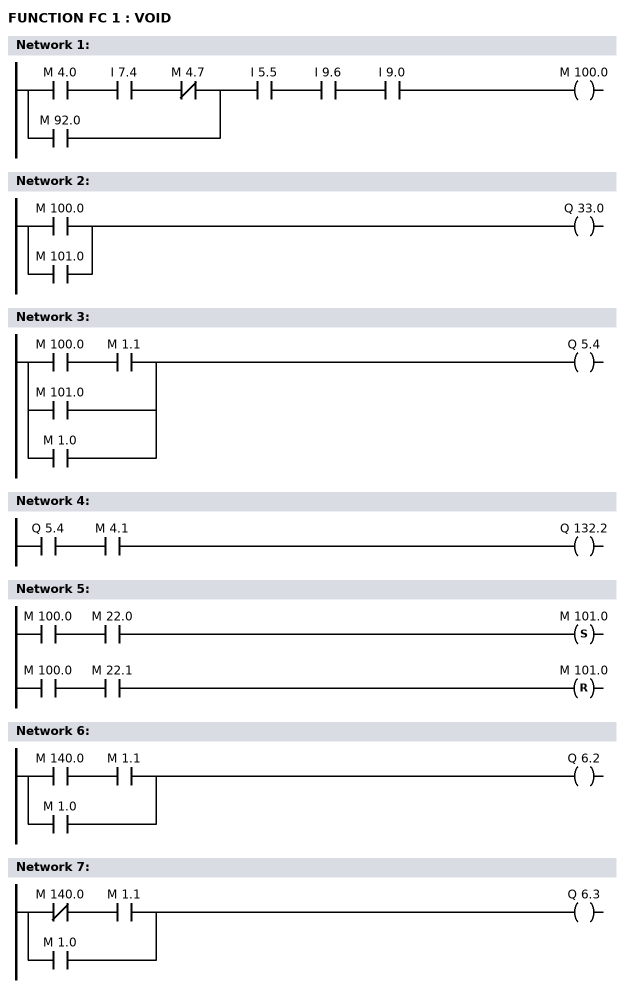

      A(    ;
      A     M      4.0;
      A     I      7.4;
      AN    M      4.7;
      O     M     92.0;
      )     ;
      A     I      5.5;
      A     I      9.6;
      A     I      9.0;
      =     M    100.0;
NETWORK
TITLE =

      O     M    100.0;
      O     M    101.0;
      =     Q     33.0;
NETWORK
TITLE =

      A     M    100.0;
      A     M      1.1;
      O     M    101.0;
      O     M      1.0;
      =     Q      5.4;
NETWORK
TITLE =

      A     Q      5.4;
      A     M      4.1;
      =     Q    132.2;
NETWORK
TITLE =

      A     M    100.0;
      A     M     22.0;
      S     M    101.0;
      A     M    100.0;
      A     M     22.1;
      R     M    101.0;
      NOP   0;
NETWORK
TITLE =

      A     M    140.0;
      A     M      1.1;
      O     M      1.0;
      =     Q      6.2;
NETWORK
TITLE =

      AN    M    140.0;
      A     M      1.1;
      O     M      1.0;
      =     Q      6.3;
NETWORK
TITLE =

      A(    ;
      A     I      8.2;
      L     S5T#150MS;
      SD    T     58;
      NOP   0;
      NOP   0;
      NOP   0;
      A     T     58;
      )     ;
      NOT   ;
      =     Q      7.5;
NETWORK
TITLE =

      A(    ;
      A     I      8.1;
      L     S5T#150MS;
      SD    T     59;
      NOP   0;
      NOP   0;
      NOP   0;
      A     T     59;
      )     ;
      NOT   ;
      =     Q      7.4;
NETWORK
TITLE =
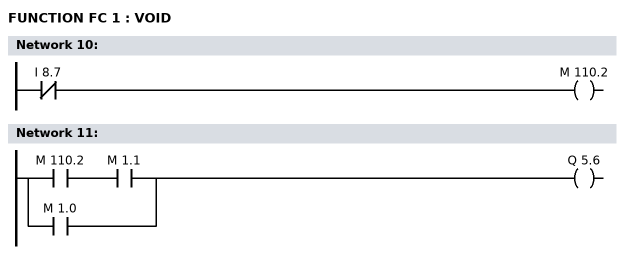

      AN    I      8.7;
      =     M    110.2;
NETWORK
TITLE =

      A     M    110.2;
      A     M      1.1;
      O     M      1.0;
      =     Q      5.6;
NETWORK
TITLE =

      O(    ;
      A     I      8.0;
      L     S5T#150MS;
      SD    T     50;
      NOP   0;
      NOP   0;
      NOP   0;
      A     T     50;
      )     ;
      O     M      1.0;
      =     Q      5.0;
NETWORK
TITLE =
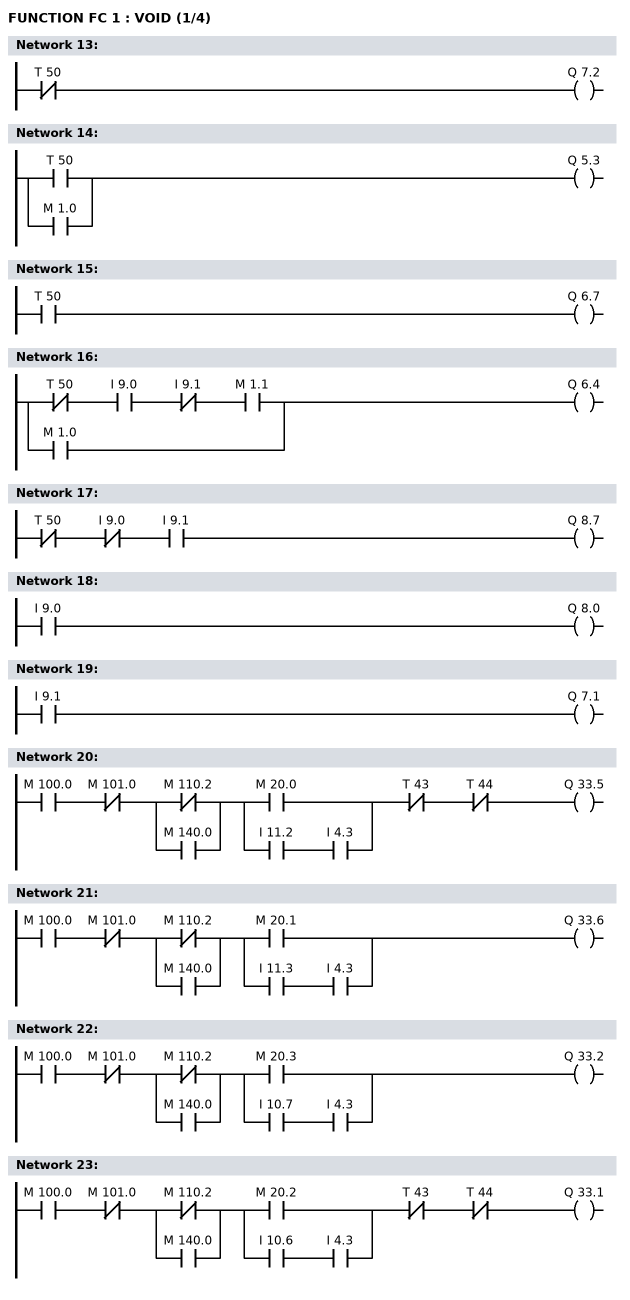

      AN    T     50;
      =     Q      7.2;
NETWORK
TITLE =

      O     T     50;
      O     M      1.0;
      =     Q      5.3;
NETWORK
TITLE =

      A     T     50;
      =     Q      6.7;
NETWORK
TITLE =

      AN    T     50;
      A     I      9.0;
      AN    I      9.1;
      A     M      1.1;
      O     M      1.0;
      =     Q      6.4;
NETWORK
TITLE =

      AN    T     50;
      AN    I      9.0;
      A     I      9.1;
      =     Q      8.7;
NETWORK
TITLE =

      A     I      9.0;
      =     Q      8.0;
NETWORK
TITLE =

      A     I      9.1;
      =     Q      7.1;
NETWORK
TITLE =

      A     M    100.0;
      AN    M    101.0;
      A(    ;
      ON    M    110.2;
      O     M    140.0;
      )     ;
      A(    ;
      O     M     20.0;
      O     ;
      A     I     11.2;
      A     I      4.3;
      )     ;
      AN    T     43;
      AN    T     44;
      =     Q     33.5;
NETWORK
TITLE =

      A     M    100.0;
      AN    M    101.0;
      A(    ;
      ON    M    110.2;
      O     M    140.0;
      )     ;
      A(    ;
      O     M     20.1;
      O     ;
      A     I     11.3;
      A     I      4.3;
      )     ;
      =     Q     33.6;
NETWORK
TITLE =

      A     M    100.0;
      AN    M    101.0;
      A(    ;
      ON    M    110.2;
      O     M    140.0;
      )     ;
      A(    ;
      O     M     20.3;
      O     ;
      A     I     10.7;
      A     I      4.3;
      )     ;
      =     Q     33.2;
NETWORK
TITLE =

      A     M    100.0;
      AN    M    101.0;
      A(    ;
      ON    M    110.2;
      O     M    140.0;
      )     ;
      A(    ;
      O     M     20.2;
      O     ;
      A     I     10.6;
      A     I      4.3;
      )     ;
      AN    T     43;
      AN    T     44;
      =     Q     33.1;
NETWORK
TITLE =
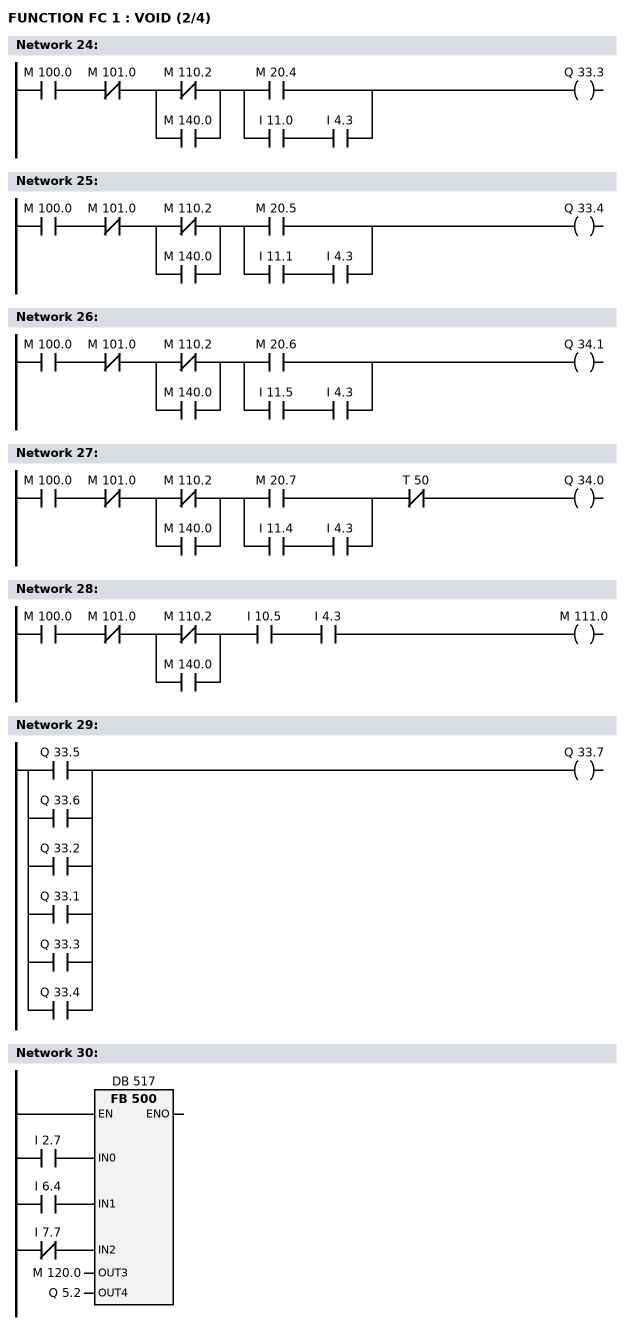

      A     M    100.0;
      AN    M    101.0;
      A(    ;
      ON    M    110.2;
      O     M    140.0;
      )     ;
      A(    ;
      O     M     20.4;
      O     ;
      A     I     11.0;
      A     I      4.3;
      )     ;
      =     Q     33.3;
NETWORK
TITLE =

      A     M    100.0;
      AN    M    101.0;
      A(    ;
      ON    M    110.2;
      O     M    140.0;
      )     ;
      A(    ;
      O     M     20.5;
      O     ;
      A     I     11.1;
      A     I      4.3;
      )     ;
      =     Q     33.4;
NETWORK
TITLE =

      A     M    100.0;
      AN    M    101.0;
      A(    ;
      ON    M    110.2;
      O     M    140.0;
      )     ;
      A(    ;
      O     M     20.6;
      O     ;
      A     I     11.5;
      A     I      4.3;
      )     ;
      =     Q     34.1;
NETWORK
TITLE =

      A     M    100.0;
      AN    M    101.0;
      A(    ;
      ON    M    110.2;
      O     M    140.0;
      )     ;
      A(    ;
      O     M     20.7;
      O     ;
      A     I     11.4;
      A     I      4.3;
      )     ;
      AN    T     50;
      =     Q     34.0;
NETWORK
TITLE =

      A     M    100.0;
      AN    M    101.0;
      A(    ;
      ON    M    110.2;
      O     M    140.0;
      )     ;
      A     I     10.5;
      A     I      4.3;
      =     M    111.0;
NETWORK
TITLE =

      O     Q     33.5;
      O     Q     33.6;
      O     Q     33.2;
      O     Q     33.1;
      O     Q     33.3;
      O     Q     33.4;
      =     Q     33.7;
NETWORK
TITLE =

      A     I      2.7;
      =     L      0.0;
      BLD   103;
      A     I      6.4;
      =     L      0.1;
      BLD   103;
      AN    I      7.7;
      =     L      0.2;
      BLD   103;
      CALL FB   500 , DB   517 (
           IN0                      := L      0.0,
           IN1                      := L      0.1,
           IN2                      := L      0.2,
           OUT3                     := M    120.0,
           OUT4                     := Q      5.2);
      NOP   0;
NETWORK
TITLE =
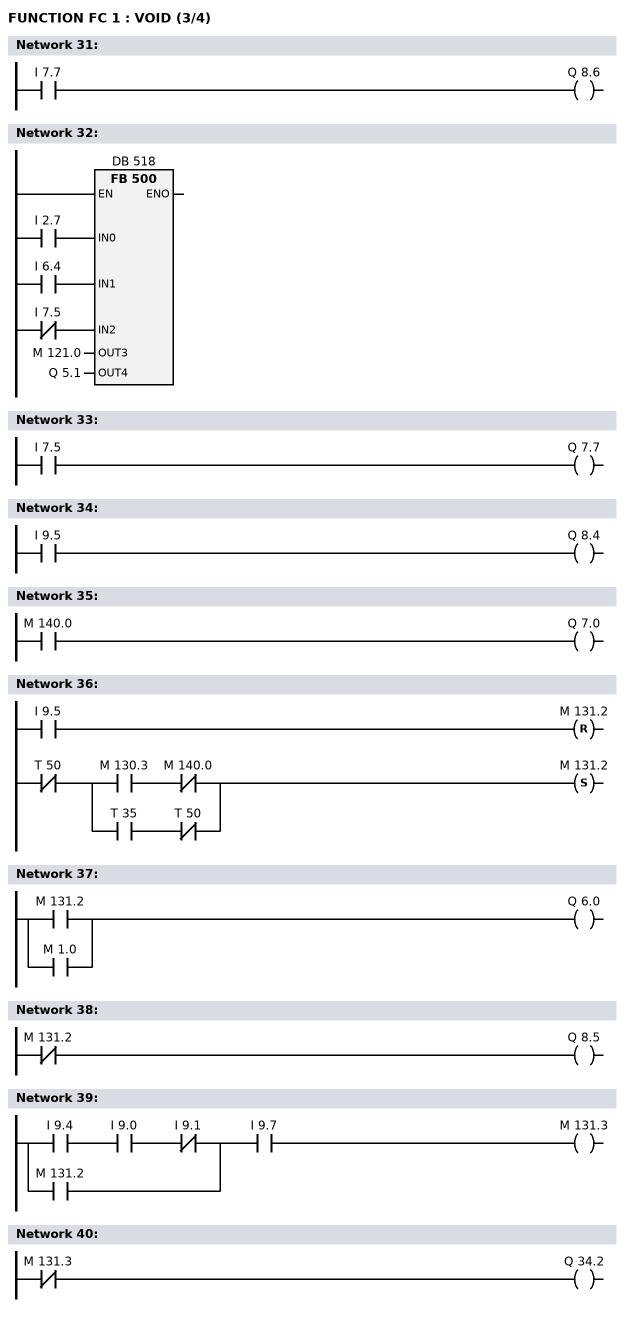

      A     I      7.7;
      =     Q      8.6;
NETWORK
TITLE =

      A     I      2.7;
      =     L      0.0;
      BLD   103;
      A     I      6.4;
      =     L      0.1;
      BLD   103;
      AN    I      7.5;
      =     L      0.2;
      BLD   103;
      CALL FB   500 , DB   518 (
           IN0                      := L      0.0,
           IN1                      := L      0.1,
           IN2                      := L      0.2,
           OUT3                     := M    121.0,
           OUT4                     := Q      5.1);
      NOP   0;
NETWORK
TITLE =

      A     I      7.5;
      =     Q      7.7;
NETWORK
TITLE =

      A     I      9.5;
      =     Q      8.4;
NETWORK
TITLE =

      A     M    140.0;
      =     Q      7.0;
NETWORK
TITLE =

      A     I      9.5;
      R     M    131.2;
      AN    T     50;
      A(    ;
      A     M    130.3;
      AN    M    140.0;
      O     ;
      A     T     35;
      AN    T     50;
      )     ;
      S     M    131.2;
      NOP   0;
NETWORK
TITLE =

      O     M    131.2;
      O     M      1.0;
      =     Q      6.0;
NETWORK
TITLE =

      AN    M    131.2;
      =     Q      8.5;
NETWORK
TITLE =

      A(    ;
      A     I      9.4;
      A     I      9.0;
      AN    I      9.1;
      O     M    131.2;
      )     ;
      A     I      9.7;
      =     M    131.3;
NETWORK
TITLE =

      AN    M    131.3;
      =     Q     34.2;
NETWORK
TITLE =
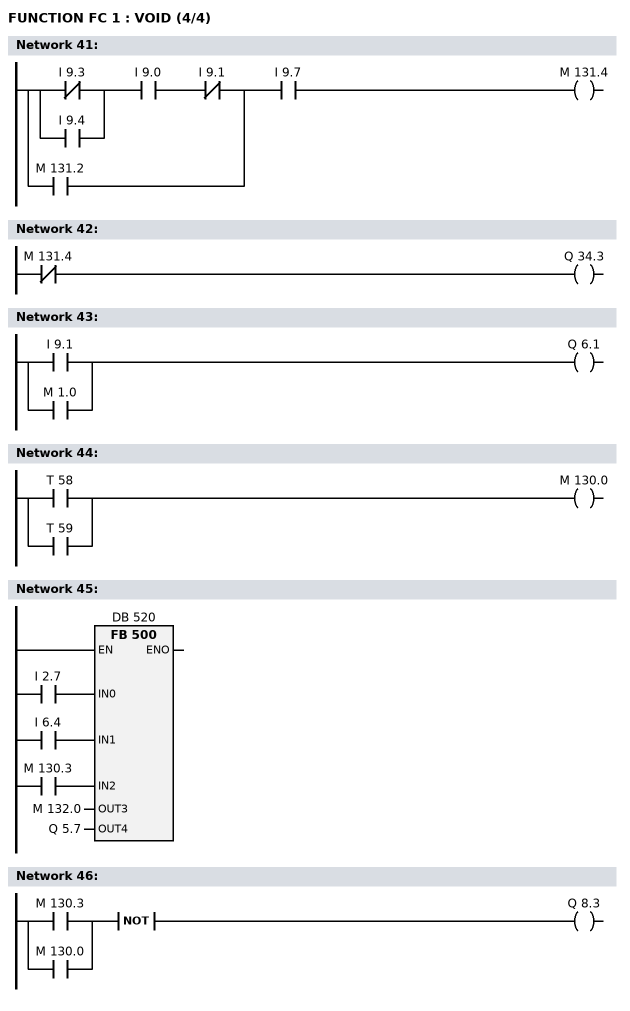

      A(    ;
      A(    ;
      ON    I      9.3;
      O     I      9.4;
      )     ;
      A     I      9.0;
      AN    I      9.1;
      O     M    131.2;
      )     ;
      A     I      9.7;
      =     M    131.4;
NETWORK
TITLE =

      AN    M    131.4;
      =     Q     34.3;
NETWORK
TITLE =

      O     I      9.1;
      O     M      1.0;
      =     Q      6.1;
NETWORK
TITLE =

      O     T     58;
      O     T     59;
      =     M    130.0;
NETWORK
TITLE =

      A     I      2.7;
      =     L      0.0;
      BLD   103;
      A     I      6.4;
      =     L      0.1;
      BLD   103;
      A     M    130.3;
      =     L      0.2;
      BLD   103;
      CALL FB   500 , DB   520 (
           IN0                      := L      0.0,
           IN1                      := L      0.1,
           IN2                      := L      0.2,
           OUT3                     := M    132.0,
           OUT4                     := Q      5.7);
      NOP   0;
NETWORK
TITLE =

      A(    ;
      O     M    130.3;
      O     M    130.0;
      )     ;
      NOT   ;
      =     Q      8.3;
NETWORK
TITLE =

      A(    ;
      A     I      8.4;
      L     S5T#150MS;
      SD    T     43;
      NOP   0;
      NOP   0;
      NOP   0;
      A     T     43;
      )     ;
      NOT   ;
      =     Q      6.6;
NETWORK
TITLE =

      A(    ;
      A     I      8.6;
      L     S5T#150MS;
      SD    T     44;
      NOP   0;
      NOP   0;
      NOP   0;
      A     T     44;
      )     ;
      NOT   ;
      =     Q      8.1;
NETWORK
TITLE =

      A(    ;
      A     I      8.5;
      L     S5T#150MS;
      SD    T     46;
      NOP   0;
      NOP   0;
      NOP   0;
      A     T     46;
      )     ;
      NOT   ;
      =     Q      7.6;
NETWORK
TITLE =

      A(    ;
      A     I      8.3;
      L     S5T#150MS;
      SD    T     47;
      NOP   0;
      NOP   0;
      NOP   0;
      A     T     47;
      )     ;
      NOT   ;
      =     Q      8.2;
NETWORK
TITLE =
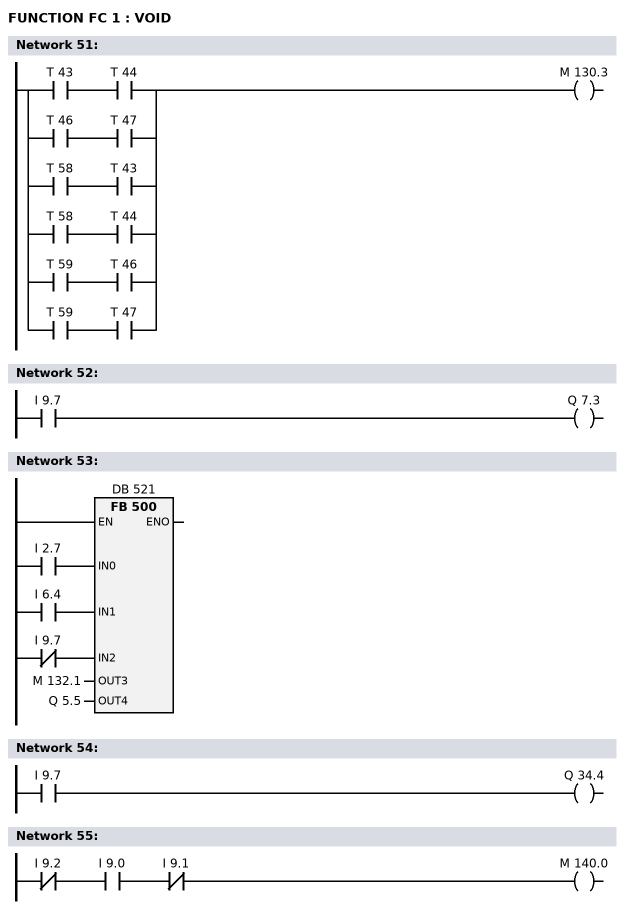

      A     T     43;
      A     T     44;
      O     ;
      A     T     46;
      A     T     47;
      O     ;
      A     T     58;
      A     T     43;
      O     ;
      A     T     58;
      A     T     44;
      O     ;
      A     T     59;
      A     T     46;
      O     ;
      A     T     59;
      A     T     47;
      =     M    130.3;
NETWORK
TITLE =

      A     I      9.7;
      =     Q      7.3;
NETWORK
TITLE =

      A     I      2.7;
      =     L      0.0;
      BLD   103;
      A     I      6.4;
      =     L      0.1;
      BLD   103;
      AN    I      9.7;
      =     L      0.2;
      BLD   103;
      CALL FB   500 , DB   521 (
           IN0                      := L      0.0,
           IN1                      := L      0.1,
           IN2                      := L      0.2,
           OUT3                     := M    132.1,
           OUT4                     := Q      5.5);
      NOP   0;
NETWORK
TITLE =

      A     I      9.7;
      =     Q     34.4;
NETWORK
TITLE =

      AN    I      9.2;
      A     I      9.0;
      AN    I      9.1;
      =     M    140.0;
END_FUNCTION

FUNCTION FC 2 : VOID
VERSION : 0.1

BEGIN
NETWORK
TITLE =
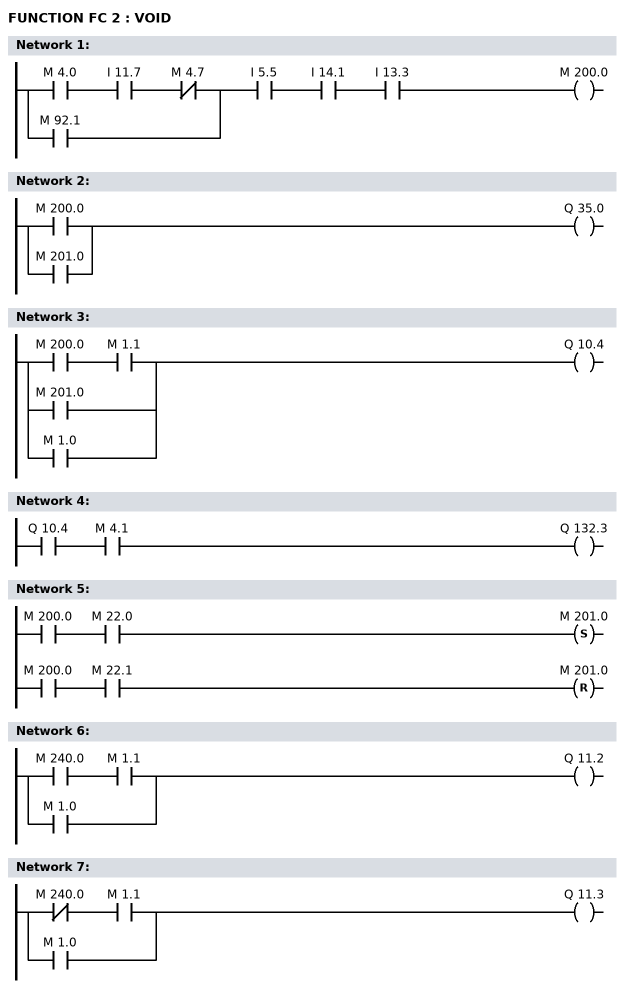

      A(    ;
      A     M      4.0;
      A     I     11.7;
      AN    M      4.7;
      O     M     92.1;
      )     ;
      A     I      5.5;
      A     I     14.1;
      A     I     13.3;
      =     M    200.0;
NETWORK
TITLE =

      O     M    200.0;
      O     M    201.0;
      =     Q     35.0;
NETWORK
TITLE =

      A     M    200.0;
      A     M      1.1;
      O     M    201.0;
      O     M      1.0;
      =     Q     10.4;
NETWORK
TITLE =

      A     Q     10.4;
      A     M      4.1;
      =     Q    132.3;
NETWORK
TITLE =

      A     M    200.0;
      A     M     22.0;
      S     M    201.0;
      A     M    200.0;
      A     M     22.1;
      R     M    201.0;
      NOP   0;
NETWORK
TITLE =

      A     M    240.0;
      A     M      1.1;
      O     M      1.0;
      =     Q     11.2;
NETWORK
TITLE =

      AN    M    240.0;
      A     M      1.1;
      O     M      1.0;
      =     Q     11.3;
NETWORK
TITLE =

      A(    ;
      A     I     12.5;
      L     S5T#150MS;
      SD    T     78;
      NOP   0;
      NOP   0;
      NOP   0;
      A     T     78;
      )     ;
      NOT   ;
      =     Q     12.5;
NETWORK
TITLE =

      A(    ;
      A     I     12.4;
      L     S5T#150MS;
      SD    T     79;
      NOP   0;
      NOP   0;
      NOP   0;
      A     T     79;
      )     ;
      NOT   ;
      =     Q     12.4;
NETWORK
TITLE =
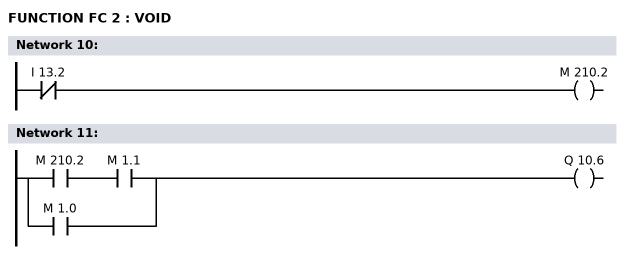

      AN    I     13.2;
      =     M    210.2;
NETWORK
TITLE =

      A     M    210.2;
      A     M      1.1;
      O     M      1.0;
      =     Q     10.6;
NETWORK
TITLE =

      O(    ;
      A     I     12.3;
      L     S5T#150MS;
      SD    T     70;
      NOP   0;
      NOP   0;
      NOP   0;
      A     T     70;
      )     ;
      O     M      1.0;
      =     Q     10.0;
NETWORK
TITLE =
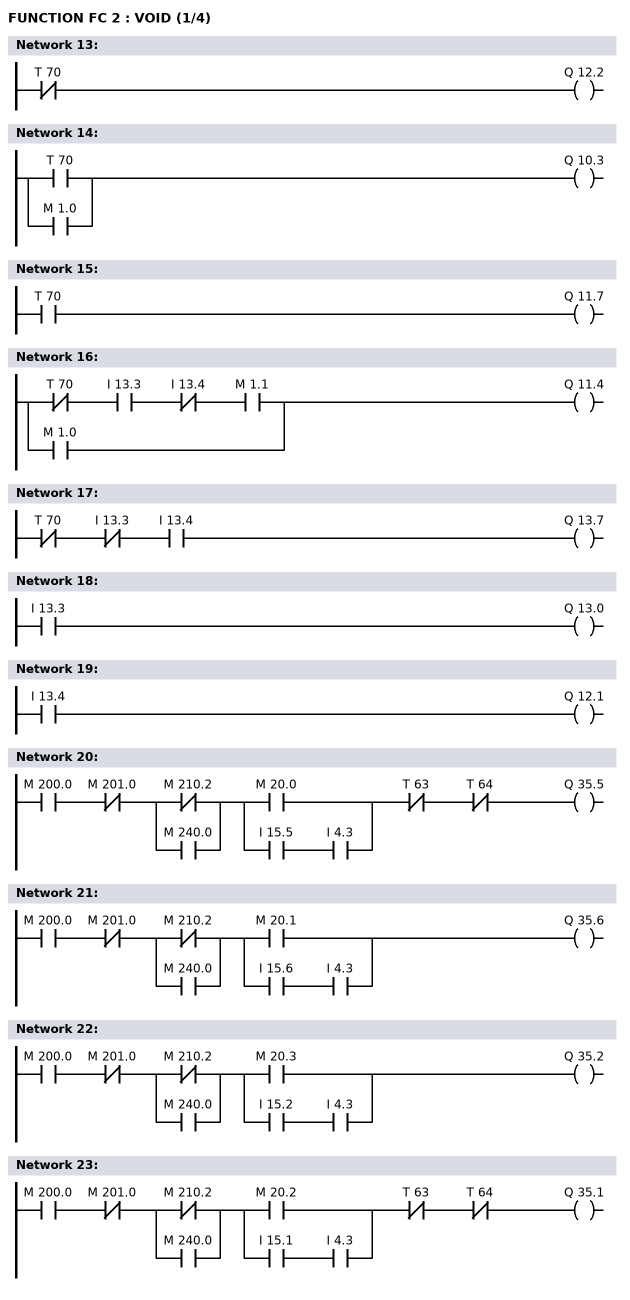

      AN    T     70;
      =     Q     12.2;
NETWORK
TITLE =

      O     T     70;
      O     M      1.0;
      =     Q     10.3;
NETWORK
TITLE =

      A     T     70;
      =     Q     11.7;
NETWORK
TITLE =

      AN    T     70;
      A     I     13.3;
      AN    I     13.4;
      A     M      1.1;
      O     M      1.0;
      =     Q     11.4;
NETWORK
TITLE =

      AN    T     70;
      AN    I     13.3;
      A     I     13.4;
      =     Q     13.7;
NETWORK
TITLE =

      A     I     13.3;
      =     Q     13.0;
NETWORK
TITLE =

      A     I     13.4;
      =     Q     12.1;
NETWORK
TITLE =

      A     M    200.0;
      AN    M    201.0;
      A(    ;
      ON    M    210.2;
      O     M    240.0;
      )     ;
      A(    ;
      O     M     20.0;
      O     ;
      A     I     15.5;
      A     I      4.3;
      )     ;
      AN    T     63;
      AN    T     64;
      =     Q     35.5;
NETWORK
TITLE =

      A     M    200.0;
      AN    M    201.0;
      A(    ;
      ON    M    210.2;
      O     M    240.0;
      )     ;
      A(    ;
      O     M     20.1;
      O     ;
      A     I     15.6;
      A     I      4.3;
      )     ;
      =     Q     35.6;
NETWORK
TITLE =

      A     M    200.0;
      AN    M    201.0;
      A(    ;
      ON    M    210.2;
      O     M    240.0;
      )     ;
      A(    ;
      O     M     20.3;
      O     ;
      A     I     15.2;
      A     I      4.3;
      )     ;
      =     Q     35.2;
NETWORK
TITLE =

      A     M    200.0;
      AN    M    201.0;
      A(    ;
      ON    M    210.2;
      O     M    240.0;
      )     ;
      A(    ;
      O     M     20.2;
      O     ;
      A     I     15.1;
      A     I      4.3;
      )     ;
      AN    T     63;
      AN    T     64;
      =     Q     35.1;
NETWORK
TITLE =
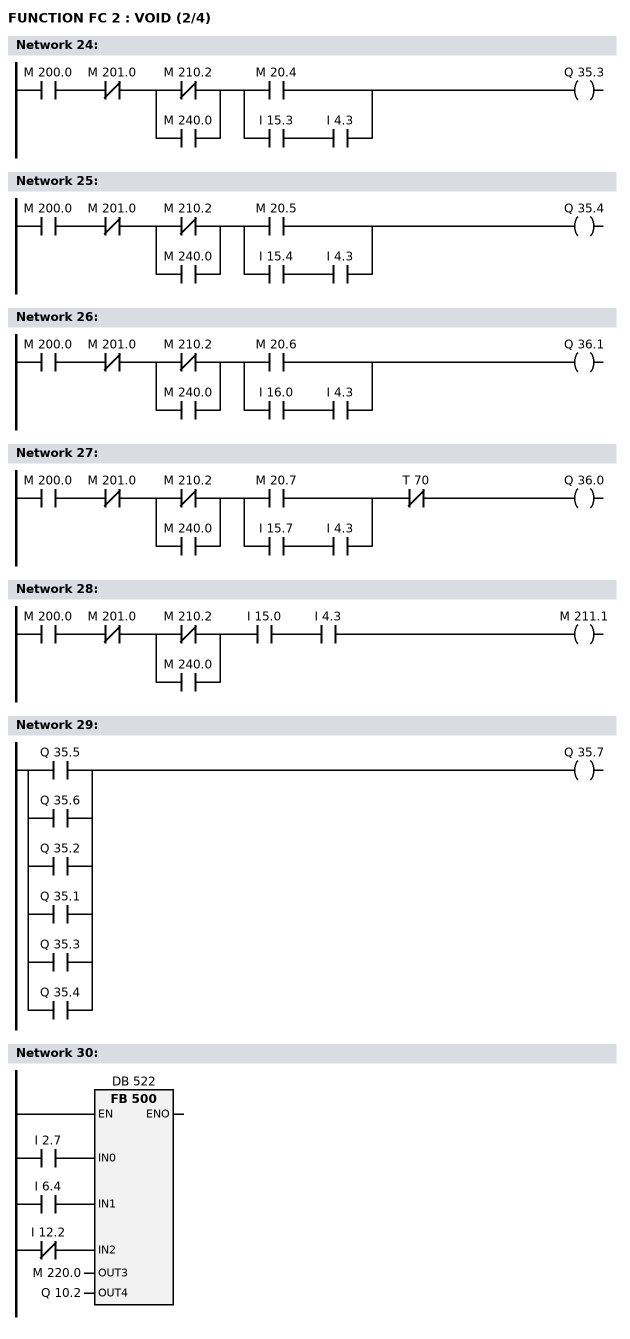

      A     M    200.0;
      AN    M    201.0;
      A(    ;
      ON    M    210.2;
      O     M    240.0;
      )     ;
      A(    ;
      O     M     20.4;
      O     ;
      A     I     15.3;
      A     I      4.3;
      )     ;
      =     Q     35.3;
NETWORK
TITLE =

      A     M    200.0;
      AN    M    201.0;
      A(    ;
      ON    M    210.2;
      O     M    240.0;
      )     ;
      A(    ;
      O     M     20.5;
      O     ;
      A     I     15.4;
      A     I      4.3;
      )     ;
      =     Q     35.4;
NETWORK
TITLE =

      A     M    200.0;
      AN    M    201.0;
      A(    ;
      ON    M    210.2;
      O     M    240.0;
      )     ;
      A(    ;
      O     M     20.6;
      O     ;
      A     I     16.0;
      A     I      4.3;
      )     ;
      =     Q     36.1;
NETWORK
TITLE =

      A     M    200.0;
      AN    M    201.0;
      A(    ;
      ON    M    210.2;
      O     M    240.0;
      )     ;
      A(    ;
      O     M     20.7;
      O     ;
      A     I     15.7;
      A     I      4.3;
      )     ;
      AN    T     70;
      =     Q     36.0;
NETWORK
TITLE =

      A     M    200.0;
      AN    M    201.0;
      A(    ;
      ON    M    210.2;
      O     M    240.0;
      )     ;
      A     I     15.0;
      A     I      4.3;
      =     M    211.1;
NETWORK
TITLE =

      O     Q     35.5;
      O     Q     35.6;
      O     Q     35.2;
      O     Q     35.1;
      O     Q     35.3;
      O     Q     35.4;
      =     Q     35.7;
NETWORK
TITLE =

      A     I      2.7;
      =     L      0.0;
      BLD   103;
      A     I      6.4;
      =     L      0.1;
      BLD   103;
      AN    I     12.2;
      =     L      0.2;
      BLD   103;
      CALL FB   500 , DB   522 (
           IN0                      := L      0.0,
           IN1                      := L      0.1,
           IN2                      := L      0.2,
           OUT3                     := M    220.0,
           OUT4                     := Q     10.2);
      NOP   0;
NETWORK
TITLE =
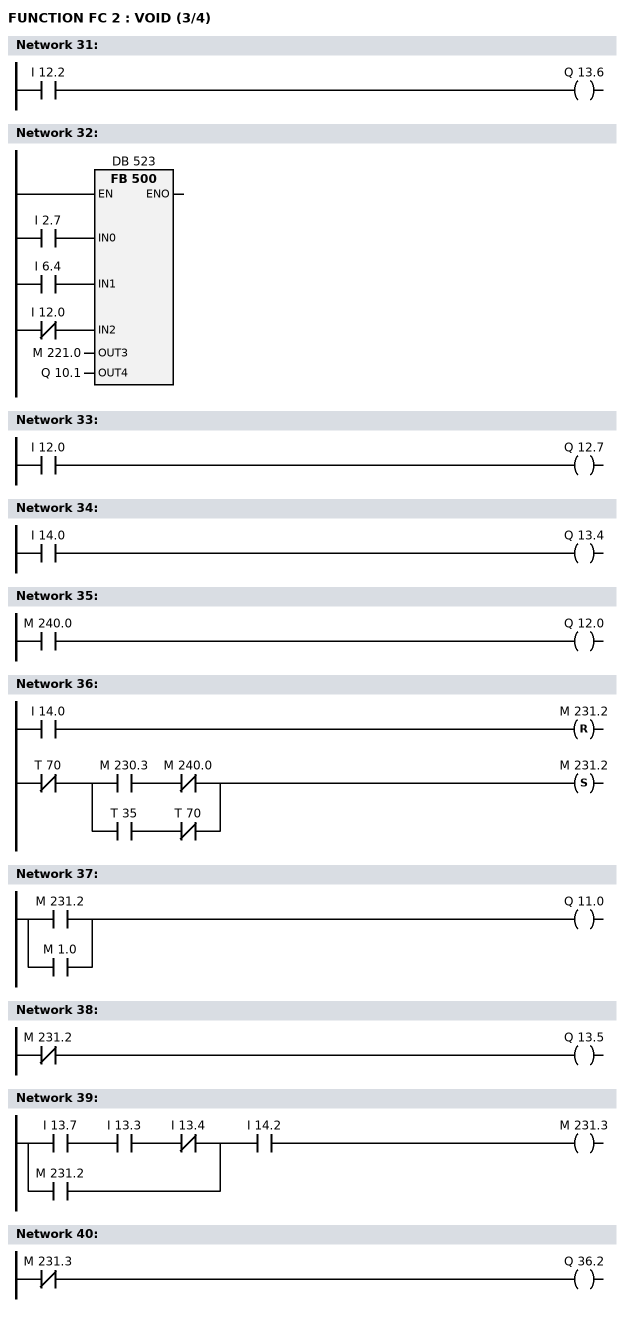

      A     I     12.2;
      =     Q     13.6;
NETWORK
TITLE =

      A     I      2.7;
      =     L      0.0;
      BLD   103;
      A     I      6.4;
      =     L      0.1;
      BLD   103;
      AN    I     12.0;
      =     L      0.2;
      BLD   103;
      CALL FB   500 , DB   523 (
           IN0                      := L      0.0,
           IN1                      := L      0.1,
           IN2                      := L      0.2,
           OUT3                     := M    221.0,
           OUT4                     := Q     10.1);
      NOP   0;
NETWORK
TITLE =

      A     I     12.0;
      =     Q     12.7;
NETWORK
TITLE =

      A     I     14.0;
      =     Q     13.4;
NETWORK
TITLE =

      A     M    240.0;
      =     Q     12.0;
NETWORK
TITLE =

      A     I     14.0;
      R     M    231.2;
      AN    T     70;
      A(    ;
      A     M    230.3;
      AN    M    240.0;
      O     ;
      A     T     35;
      AN    T     70;
      )     ;
      S     M    231.2;
      NOP   0;
NETWORK
TITLE =

      O     M    231.2;
      O     M      1.0;
      =     Q     11.0;
NETWORK
TITLE =

      AN    M    231.2;
      =     Q     13.5;
NETWORK
TITLE =

      A(    ;
      A     I     13.7;
      A     I     13.3;
      AN    I     13.4;
      O     M    231.2;
      )     ;
      A     I     14.2;
      =     M    231.3;
NETWORK
TITLE =

      AN    M    231.3;
      =     Q     36.2;
NETWORK
TITLE =
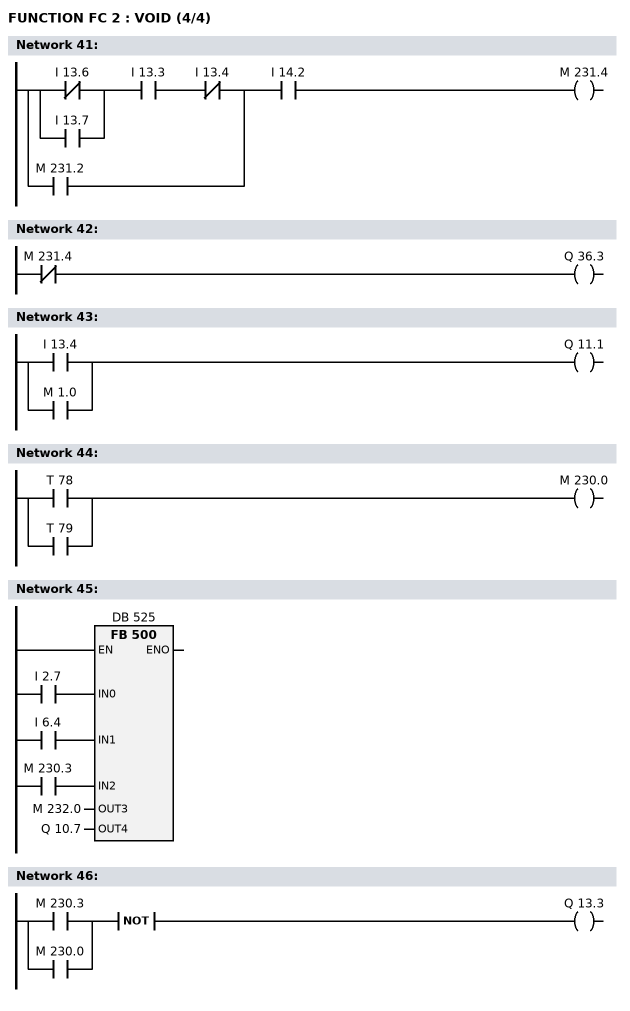

      A(    ;
      A(    ;
      ON    I     13.6;
      O     I     13.7;
      )     ;
      A     I     13.3;
      AN    I     13.4;
      O     M    231.2;
      )     ;
      A     I     14.2;
      =     M    231.4;
NETWORK
TITLE =

      AN    M    231.4;
      =     Q     36.3;
NETWORK
TITLE =

      O     I     13.4;
      O     M      1.0;
      =     Q     11.1;
NETWORK
TITLE =

      O     T     78;
      O     T     79;
      =     M    230.0;
NETWORK
TITLE =

      A     I      2.7;
      =     L      0.0;
      BLD   103;
      A     I      6.4;
      =     L      0.1;
      BLD   103;
      A     M    230.3;
      =     L      0.2;
      BLD   103;
      CALL FB   500 , DB   525 (
           IN0                      := L      0.0,
           IN1                      := L      0.1,
           IN2                      := L      0.2,
           OUT3                     := M    232.0,
           OUT4                     := Q     10.7);
      NOP   0;
NETWORK
TITLE =

      A(    ;
      O     M    230.3;
      O     M    230.0;
      )     ;
      NOT   ;
      =     Q     13.3;
NETWORK
TITLE =

      A(    ;
      A     I     12.7;
      L     S5T#150MS;
      SD    T     63;
      NOP   0;
      NOP   0;
      NOP   0;
      A     T     63;
      )     ;
      NOT   ;
      =     Q     11.6;
NETWORK
TITLE =

      A(    ;
      A     I     13.1;
      L     S5T#150MS;
      SD    T     64;
      NOP   0;
      NOP   0;
      NOP   0;
      A     T     64;
      )     ;
      NOT   ;
      =     Q     13.1;
NETWORK
TITLE =

      A(    ;
      A     I     13.0;
      L     S5T#150MS;
      SD    T     66;
      NOP   0;
      NOP   0;
      NOP   0;
      A     T     66;
      )     ;
      NOT   ;
      =     Q     12.6;
NETWORK
TITLE =

      A(    ;
      A     I     12.6;
      L     S5T#150MS;
      SD    T     67;
      NOP   0;
      NOP   0;
      NOP   0;
      A     T     67;
      )     ;
      NOT   ;
      =     Q     13.2;
NETWORK
TITLE =
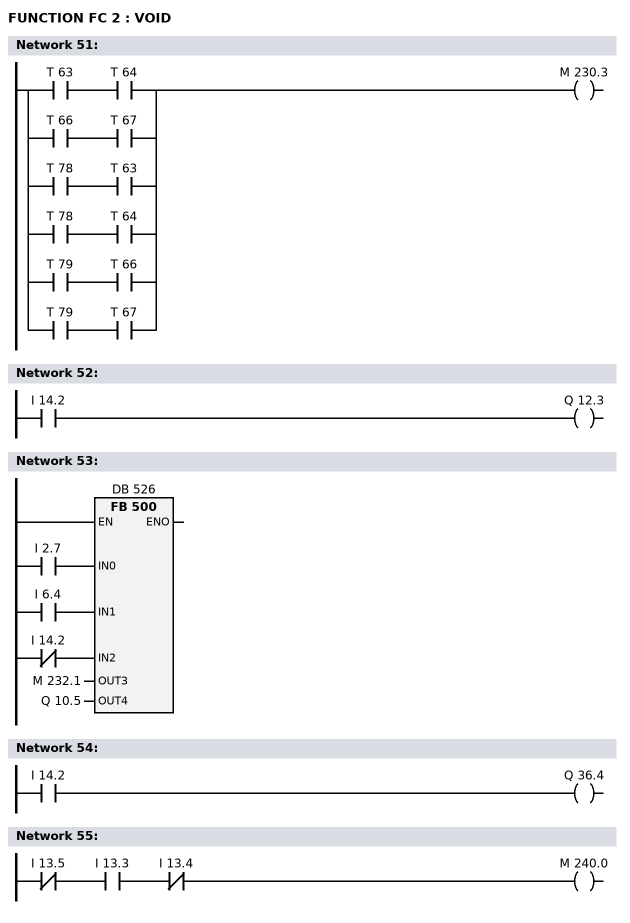

      A     T     63;
      A     T     64;
      O     ;
      A     T     66;
      A     T     67;
      O     ;
      A     T     78;
      A     T     63;
      O     ;
      A     T     78;
      A     T     64;
      O     ;
      A     T     79;
      A     T     66;
      O     ;
      A     T     79;
      A     T     67;
      =     M    230.3;
NETWORK
TITLE =

      A     I     14.2;
      =     Q     12.3;
NETWORK
TITLE =

      A     I      2.7;
      =     L      0.0;
      BLD   103;
      A     I      6.4;
      =     L      0.1;
      BLD   103;
      AN    I     14.2;
      =     L      0.2;
      BLD   103;
      CALL FB   500 , DB   526 (
           IN0                      := L      0.0,
           IN1                      := L      0.1,
           IN2                      := L      0.2,
           OUT3                     := M    232.1,
           OUT4                     := Q     10.5);
      NOP   0;
NETWORK
TITLE =

      A     I     14.2;
      =     Q     36.4;
NETWORK
TITLE =

      AN    I     13.5;
      A     I     13.3;
      AN    I     13.4;
      =     M    240.0;
END_FUNCTION

FUNCTION FC 3 : VOID
VERSION : 0.1

BEGIN
NETWORK
TITLE =
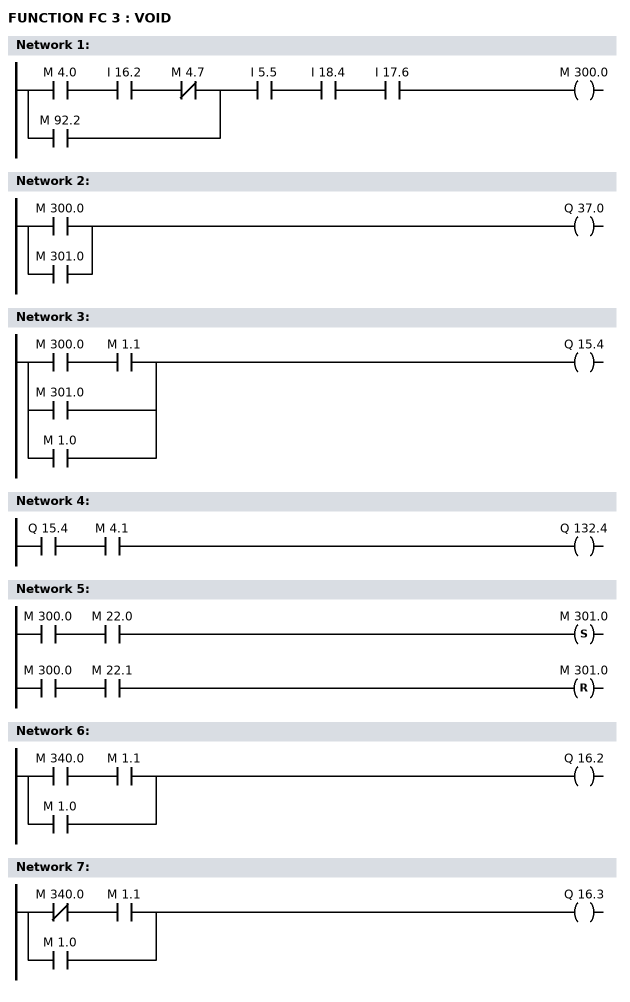

      A(    ;
      A     M      4.0;
      A     I     16.2;
      AN    M      4.7;
      O     M     92.2;
      )     ;
      A     I      5.5;
      A     I     18.4;
      A     I     17.6;
      =     M    300.0;
NETWORK
TITLE =

      O     M    300.0;
      O     M    301.0;
      =     Q     37.0;
NETWORK
TITLE =

      A     M    300.0;
      A     M      1.1;
      O     M    301.0;
      O     M      1.0;
      =     Q     15.4;
NETWORK
TITLE =

      A     Q     15.4;
      A     M      4.1;
      =     Q    132.4;
NETWORK
TITLE =

      A     M    300.0;
      A     M     22.0;
      S     M    301.0;
      A     M    300.0;
      A     M     22.1;
      R     M    301.0;
      NOP   0;
NETWORK
TITLE =

      A     M    340.0;
      A     M      1.1;
      O     M      1.0;
      =     Q     16.2;
NETWORK
TITLE =

      AN    M    340.0;
      A     M      1.1;
      O     M      1.0;
      =     Q     16.3;
NETWORK
TITLE =

      A(    ;
      A     I     17.0;
      L     S5T#150MS;
      SD    T     98;
      NOP   0;
      NOP   0;
      NOP   0;
      A     T     98;
      )     ;
      NOT   ;
      =     Q     17.5;
NETWORK
TITLE =

      A(    ;
      A     I     16.7;
      L     S5T#150MS;
      SD    T     99;
      NOP   0;
      NOP   0;
      NOP   0;
      A     T     99;
      )     ;
      NOT   ;
      =     Q     17.4;
NETWORK
TITLE =
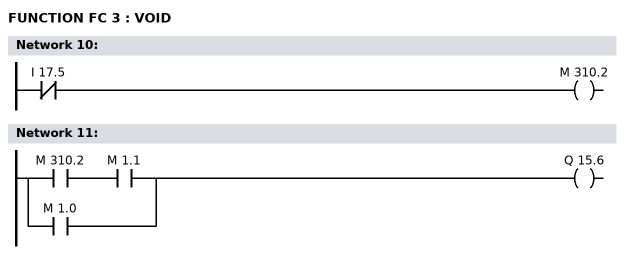

      AN    I     17.5;
      =     M    310.2;
NETWORK
TITLE =

      A     M    310.2;
      A     M      1.1;
      O     M      1.0;
      =     Q     15.6;
NETWORK
TITLE =

      O(    ;
      A     I     16.6;
      L     S5T#150MS;
      SD    T     90;
      NOP   0;
      NOP   0;
      NOP   0;
      A     T     90;
      )     ;
      O     M      1.0;
      =     Q     15.0;
NETWORK
TITLE =
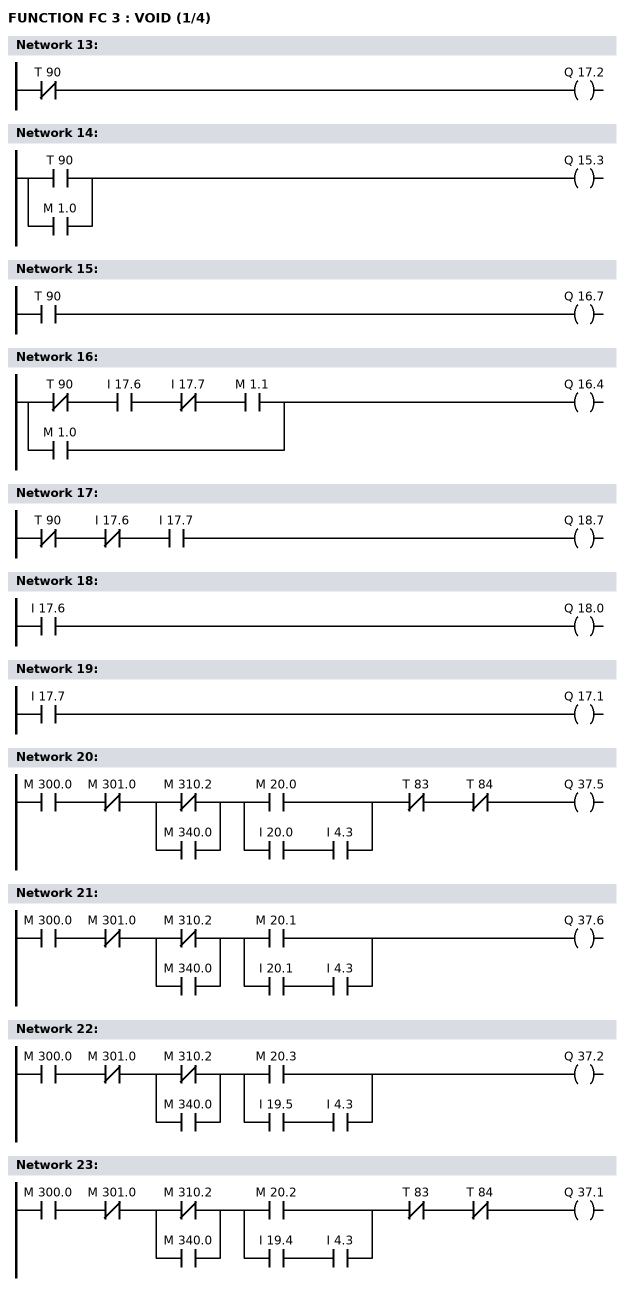

      AN    T     90;
      =     Q     17.2;
NETWORK
TITLE =

      O     T     90;
      O     M      1.0;
      =     Q     15.3;
NETWORK
TITLE =

      A     T     90;
      =     Q     16.7;
NETWORK
TITLE =

      AN    T     90;
      A     I     17.6;
      AN    I     17.7;
      A     M      1.1;
      O     M      1.0;
      =     Q     16.4;
NETWORK
TITLE =

      AN    T     90;
      AN    I     17.6;
      A     I     17.7;
      =     Q     18.7;
NETWORK
TITLE =

      A     I     17.6;
      =     Q     18.0;
NETWORK
TITLE =

      A     I     17.7;
      =     Q     17.1;
NETWORK
TITLE =

      A     M    300.0;
      AN    M    301.0;
      A(    ;
      ON    M    310.2;
      O     M    340.0;
      )     ;
      A(    ;
      O     M     20.0;
      O     ;
      A     I     20.0;
      A     I      4.3;
      )     ;
      AN    T     83;
      AN    T     84;
      =     Q     37.5;
NETWORK
TITLE =

      A     M    300.0;
      AN    M    301.0;
      A(    ;
      ON    M    310.2;
      O     M    340.0;
      )     ;
      A(    ;
      O     M     20.1;
      O     ;
      A     I     20.1;
      A     I      4.3;
      )     ;
      =     Q     37.6;
NETWORK
TITLE =

      A     M    300.0;
      AN    M    301.0;
      A(    ;
      ON    M    310.2;
      O     M    340.0;
      )     ;
      A(    ;
      O     M     20.3;
      O     ;
      A     I     19.5;
      A     I      4.3;
      )     ;
      =     Q     37.2;
NETWORK
TITLE =

      A     M    300.0;
      AN    M    301.0;
      A(    ;
      ON    M    310.2;
      O     M    340.0;
      )     ;
      A(    ;
      O     M     20.2;
      O     ;
      A     I     19.4;
      A     I      4.3;
      )     ;
      AN    T     83;
      AN    T     84;
      =     Q     37.1;
NETWORK
TITLE =
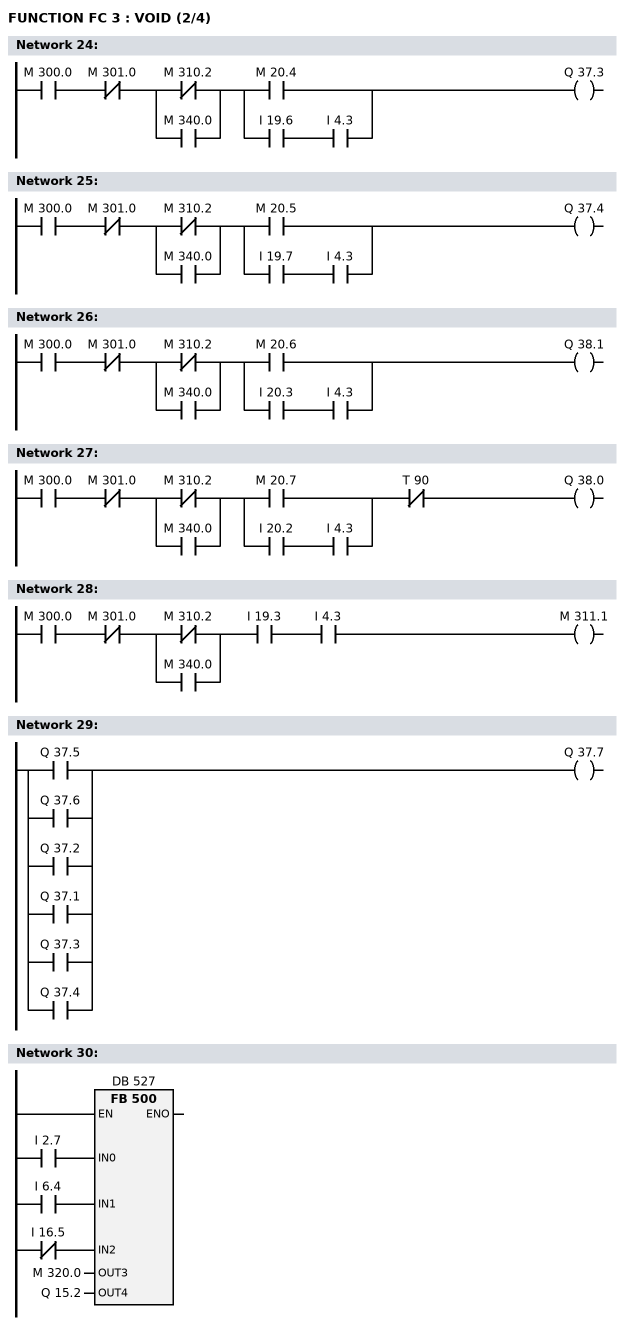

      A     M    300.0;
      AN    M    301.0;
      A(    ;
      ON    M    310.2;
      O     M    340.0;
      )     ;
      A(    ;
      O     M     20.4;
      O     ;
      A     I     19.6;
      A     I      4.3;
      )     ;
      =     Q     37.3;
NETWORK
TITLE =

      A     M    300.0;
      AN    M    301.0;
      A(    ;
      ON    M    310.2;
      O     M    340.0;
      )     ;
      A(    ;
      O     M     20.5;
      O     ;
      A     I     19.7;
      A     I      4.3;
      )     ;
      =     Q     37.4;
NETWORK
TITLE =

      A     M    300.0;
      AN    M    301.0;
      A(    ;
      ON    M    310.2;
      O     M    340.0;
      )     ;
      A(    ;
      O     M     20.6;
      O     ;
      A     I     20.3;
      A     I      4.3;
      )     ;
      =     Q     38.1;
NETWORK
TITLE =

      A     M    300.0;
      AN    M    301.0;
      A(    ;
      ON    M    310.2;
      O     M    340.0;
      )     ;
      A(    ;
      O     M     20.7;
      O     ;
      A     I     20.2;
      A     I      4.3;
      )     ;
      AN    T     90;
      =     Q     38.0;
NETWORK
TITLE =

      A     M    300.0;
      AN    M    301.0;
      A(    ;
      ON    M    310.2;
      O     M    340.0;
      )     ;
      A     I     19.3;
      A     I      4.3;
      =     M    311.1;
NETWORK
TITLE =

      O     Q     37.5;
      O     Q     37.6;
      O     Q     37.2;
      O     Q     37.1;
      O     Q     37.3;
      O     Q     37.4;
      =     Q     37.7;
NETWORK
TITLE =

      A     I      2.7;
      =     L      0.0;
      BLD   103;
      A     I      6.4;
      =     L      0.1;
      BLD   103;
      AN    I     16.5;
      =     L      0.2;
      BLD   103;
      CALL FB   500 , DB   527 (
           IN0                      := L      0.0,
           IN1                      := L      0.1,
           IN2                      := L      0.2,
           OUT3                     := M    320.0,
           OUT4                     := Q     15.2);
      NOP   0;
NETWORK
TITLE =
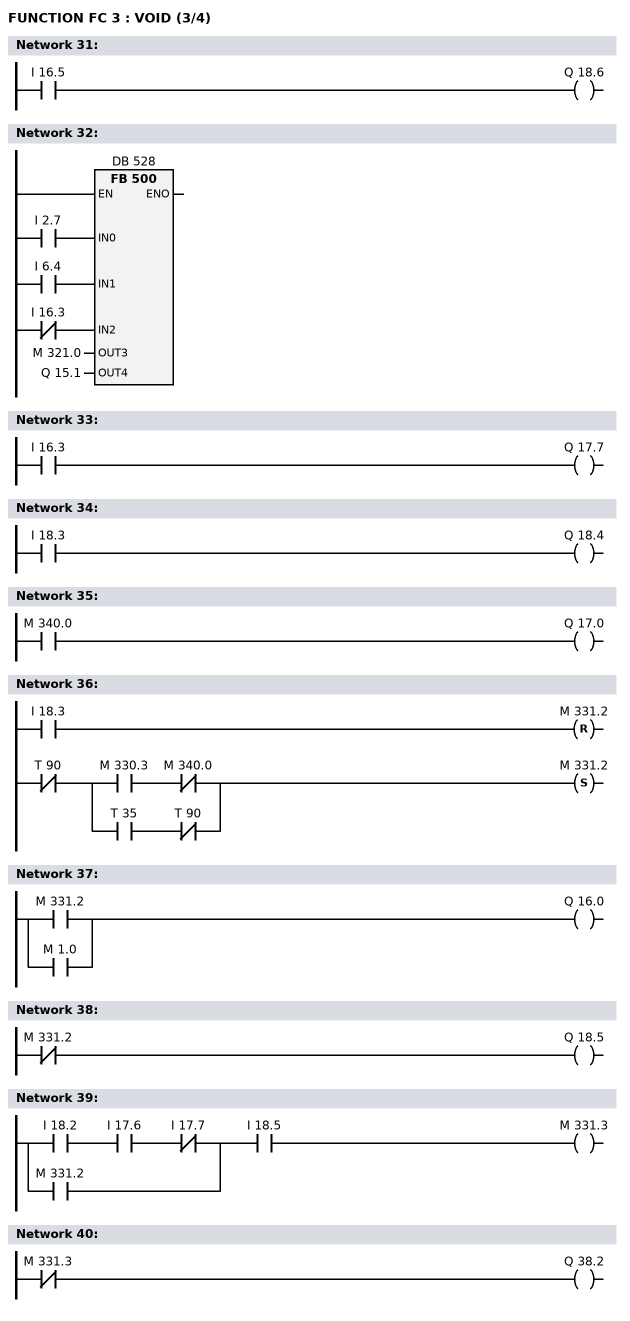

      A     I     16.5;
      =     Q     18.6;
NETWORK
TITLE =

      A     I      2.7;
      =     L      0.0;
      BLD   103;
      A     I      6.4;
      =     L      0.1;
      BLD   103;
      AN    I     16.3;
      =     L      0.2;
      BLD   103;
      CALL FB   500 , DB   528 (
           IN0                      := L      0.0,
           IN1                      := L      0.1,
           IN2                      := L      0.2,
           OUT3                     := M    321.0,
           OUT4                     := Q     15.1);
      NOP   0;
NETWORK
TITLE =

      A     I     16.3;
      =     Q     17.7;
NETWORK
TITLE =

      A     I     18.3;
      =     Q     18.4;
NETWORK
TITLE =

      A     M    340.0;
      =     Q     17.0;
NETWORK
TITLE =

      A     I     18.3;
      R     M    331.2;
      AN    T     90;
      A(    ;
      A     M    330.3;
      AN    M    340.0;
      O     ;
      A     T     35;
      AN    T     90;
      )     ;
      S     M    331.2;
      NOP   0;
NETWORK
TITLE =

      O     M    331.2;
      O     M      1.0;
      =     Q     16.0;
NETWORK
TITLE =

      AN    M    331.2;
      =     Q     18.5;
NETWORK
TITLE =

      A(    ;
      A     I     18.2;
      A     I     17.6;
      AN    I     17.7;
      O     M    331.2;
      )     ;
      A     I     18.5;
      =     M    331.3;
NETWORK
TITLE =

      AN    M    331.3;
      =     Q     38.2;
NETWORK
TITLE =
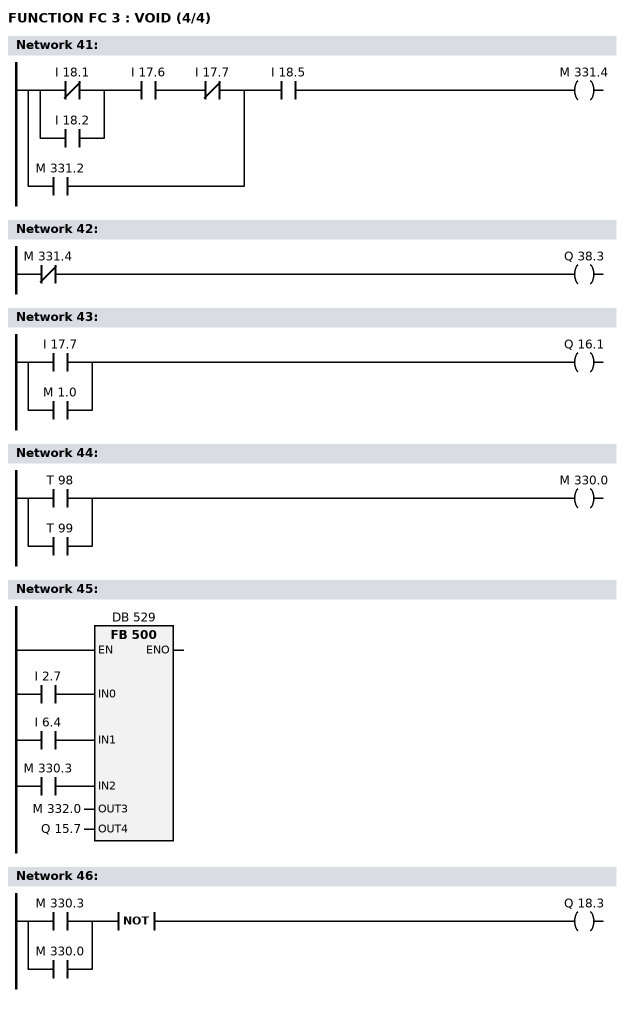

      A(    ;
      A(    ;
      ON    I     18.1;
      O     I     18.2;
      )     ;
      A     I     17.6;
      AN    I     17.7;
      O     M    331.2;
      )     ;
      A     I     18.5;
      =     M    331.4;
NETWORK
TITLE =

      AN    M    331.4;
      =     Q     38.3;
NETWORK
TITLE =

      O     I     17.7;
      O     M      1.0;
      =     Q     16.1;
NETWORK
TITLE =

      O     T     98;
      O     T     99;
      =     M    330.0;
NETWORK
TITLE =

      A     I      2.7;
      =     L      0.0;
      BLD   103;
      A     I      6.4;
      =     L      0.1;
      BLD   103;
      A     M    330.3;
      =     L      0.2;
      BLD   103;
      CALL FB   500 , DB   529 (
           IN0                      := L      0.0,
           IN1                      := L      0.1,
           IN2                      := L      0.2,
           OUT3                     := M    332.0,
           OUT4                     := Q     15.7);
      NOP   0;
NETWORK
TITLE =

      A(    ;
      O     M    330.3;
      O     M    330.0;
      )     ;
      NOT   ;
      =     Q     18.3;
NETWORK
TITLE =

      A(    ;
      A     I     17.2;
      L     S5T#150MS;
      SD    T     83;
      NOP   0;
      NOP   0;
      NOP   0;
      A     T     83;
      )     ;
      NOT   ;
      =     Q     16.6;
NETWORK
TITLE =

      A(    ;
      A     I     17.4;
      L     S5T#150MS;
      SD    T     84;
      NOP   0;
      NOP   0;
      NOP   0;
      A     T     84;
      )     ;
      NOT   ;
      =     Q     18.1;
NETWORK
TITLE =

      A(    ;
      A     I     17.3;
      L     S5T#150MS;
      SD    T     86;
      NOP   0;
      NOP   0;
      NOP   0;
      A     T     86;
      )     ;
      NOT   ;
      =     Q     17.6;
NETWORK
TITLE =

      A(    ;
      A     I     17.1;
      L     S5T#150MS;
      SD    T     87;
      NOP   0;
      NOP   0;
      NOP   0;
      A     T     87;
      )     ;
      NOT   ;
      =     Q     18.2;
NETWORK
TITLE =
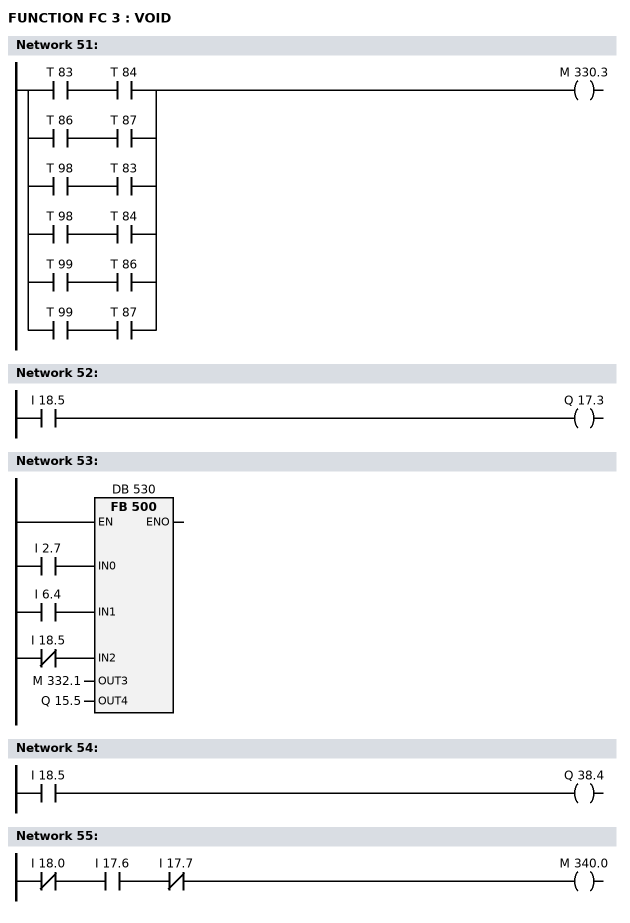

      A     T     83;
      A     T     84;
      O     ;
      A     T     86;
      A     T     87;
      O     ;
      A     T     98;
      A     T     83;
      O     ;
      A     T     98;
      A     T     84;
      O     ;
      A     T     99;
      A     T     86;
      O     ;
      A     T     99;
      A     T     87;
      =     M    330.3;
NETWORK
TITLE =

      A     I     18.5;
      =     Q     17.3;
NETWORK
TITLE =

      A     I      2.7;
      =     L      0.0;
      BLD   103;
      A     I      6.4;
      =     L      0.1;
      BLD   103;
      AN    I     18.5;
      =     L      0.2;
      BLD   103;
      CALL FB   500 , DB   530 (
           IN0                      := L      0.0,
           IN1                      := L      0.1,
           IN2                      := L      0.2,
           OUT3                     := M    332.1,
           OUT4                     := Q     15.5);
      NOP   0;
NETWORK
TITLE =

      A     I     18.5;
      =     Q     38.4;
NETWORK
TITLE =

      AN    I     18.0;
      A     I     17.6;
      AN    I     17.7;
      =     M    340.0;
END_FUNCTION

FUNCTION FC 4 : VOID
VERSION : 0.1

BEGIN
NETWORK
TITLE =
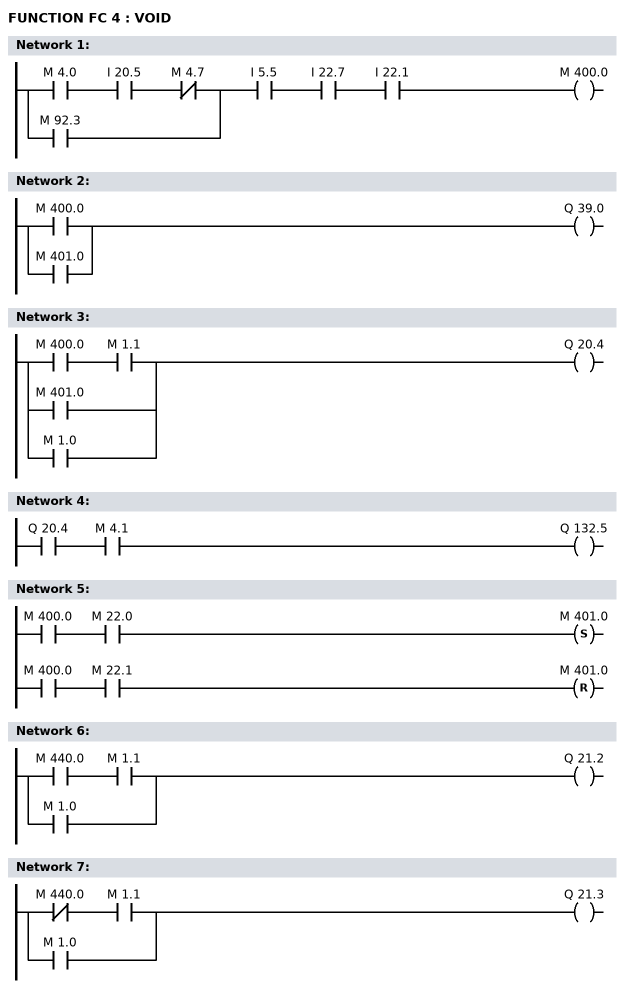

      A(    ;
      A     M      4.0;
      A     I     20.5;
      AN    M      4.7;
      O     M     92.3;
      )     ;
      A     I      5.5;
      A     I     22.7;
      A     I     22.1;
      =     M    400.0;
NETWORK
TITLE =

      O     M    400.0;
      O     M    401.0;
      =     Q     39.0;
NETWORK
TITLE =

      A     M    400.0;
      A     M      1.1;
      O     M    401.0;
      O     M      1.0;
      =     Q     20.4;
NETWORK
TITLE =

      A     Q     20.4;
      A     M      4.1;
      =     Q    132.5;
NETWORK
TITLE =

      A     M    400.0;
      A     M     22.0;
      S     M    401.0;
      A     M    400.0;
      A     M     22.1;
      R     M    401.0;
      NOP   0;
NETWORK
TITLE =

      A     M    440.0;
      A     M      1.1;
      O     M      1.0;
      =     Q     21.2;
NETWORK
TITLE =

      AN    M    440.0;
      A     M      1.1;
      O     M      1.0;
      =     Q     21.3;
NETWORK
TITLE =

      A(    ;
      A     I     21.3;
      L     S5T#150MS;
      SD    T    118;
      NOP   0;
      NOP   0;
      NOP   0;
      A     T    118;
      )     ;
      NOT   ;
      =     Q     22.5;
NETWORK
TITLE =

      A(    ;
      A     I     21.2;
      L     S5T#150MS;
      SD    T    119;
      NOP   0;
      NOP   0;
      NOP   0;
      A     T    119;
      )     ;
      NOT   ;
      =     Q     22.4;
NETWORK
TITLE =
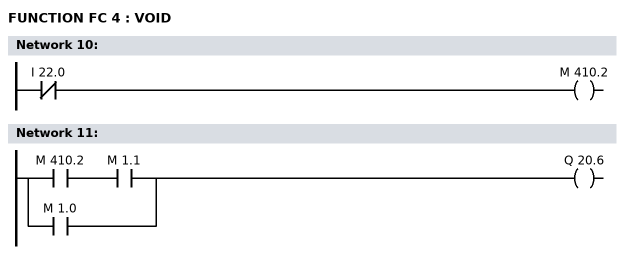

      AN    I     22.0;
      =     M    410.2;
NETWORK
TITLE =

      A     M    410.2;
      A     M      1.1;
      O     M      1.0;
      =     Q     20.6;
NETWORK
TITLE =

      O(    ;
      A     I     21.1;
      L     S5T#150MS;
      SD    T    110;
      NOP   0;
      NOP   0;
      NOP   0;
      A     T    110;
      )     ;
      O     M      1.0;
      =     Q     20.0;
NETWORK
TITLE =
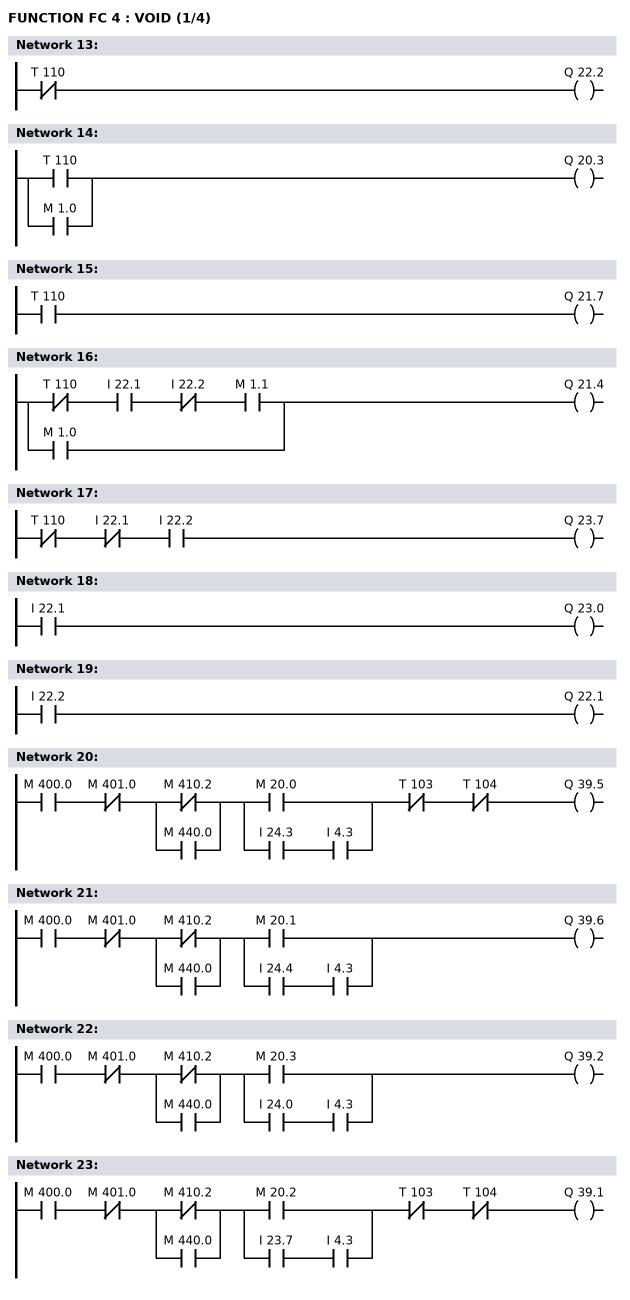

      AN    T    110;
      =     Q     22.2;
NETWORK
TITLE =

      O     T    110;
      O     M      1.0;
      =     Q     20.3;
NETWORK
TITLE =

      A     T    110;
      =     Q     21.7;
NETWORK
TITLE =

      AN    T    110;
      A     I     22.1;
      AN    I     22.2;
      A     M      1.1;
      O     M      1.0;
      =     Q     21.4;
NETWORK
TITLE =

      AN    T    110;
      AN    I     22.1;
      A     I     22.2;
      =     Q     23.7;
NETWORK
TITLE =

      A     I     22.1;
      =     Q     23.0;
NETWORK
TITLE =

      A     I     22.2;
      =     Q     22.1;
NETWORK
TITLE =

      A     M    400.0;
      AN    M    401.0;
      A(    ;
      ON    M    410.2;
      O     M    440.0;
      )     ;
      A(    ;
      O     M     20.0;
      O     ;
      A     I     24.3;
      A     I      4.3;
      )     ;
      AN    T    103;
      AN    T    104;
      =     Q     39.5;
NETWORK
TITLE =

      A     M    400.0;
      AN    M    401.0;
      A(    ;
      ON    M    410.2;
      O     M    440.0;
      )     ;
      A(    ;
      O     M     20.1;
      O     ;
      A     I     24.4;
      A     I      4.3;
      )     ;
      =     Q     39.6;
NETWORK
TITLE =

      A     M    400.0;
      AN    M    401.0;
      A(    ;
      ON    M    410.2;
      O     M    440.0;
      )     ;
      A(    ;
      O     M     20.3;
      O     ;
      A     I     24.0;
      A     I      4.3;
      )     ;
      =     Q     39.2;
NETWORK
TITLE =

      A     M    400.0;
      AN    M    401.0;
      A(    ;
      ON    M    410.2;
      O     M    440.0;
      )     ;
      A(    ;
      O     M     20.2;
      O     ;
      A     I     23.7;
      A     I      4.3;
      )     ;
      AN    T    103;
      AN    T    104;
      =     Q     39.1;
NETWORK
TITLE =
